INTERFACE I_XtsNctTool EXTENDS I_Base

PROPERTY NctBaseUnit : I_XtsNctBaseUnit
GET
END_GET
SET
END_SET
END_PROPERTY

{attribute 'monitoring' := 'call'}
PROPERTY Simulated : BOOL
GET
END_GET
SET
END_SET
END_PROPERTY

END_INTERFACE

(* stored: Version 1.1.0.1, ProductVersion 3.1.4026.21
   Itf I_XtsNctTool: Id {e66a611d-cdb3-43c9-a001-92be26719739}
   Property NctBaseUnit: Id {a2e368c0-964b-4562-85eb-16eacc5b34e7}
   Get Get: Id {953b0eb2-e7e9-41d9-9f4d-778e81783e2d}
   Set Set: Id {57b6402f-abb6-4d8b-ba84-696fa4eccedb}
   Property Simulated: Id {0aa4e837-0f99-40c8-90f8-5e262fef8547}
   Get Get: Id {0b918d6f-507b-46af-a7e1-125e19df9ce3}
   Set Set: Id {c39ce664-6e7d-493c-8286-2884394fcaa3} *)
